ADAPTER arm_sensor (* Adapter Interface *)
  (* Standard: 61499-1 *)
  (* Version 0.0, 10/22/2026, lizar, Schneider Electric *)
  PACKAGE Main;
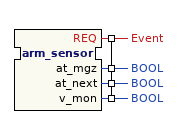
  EVENT_OUTPUT
    REQ WITH at_mgz, at_next, v_mon; (* Confirmation from Plug *)
  END_EVENT
  VAR_OUTPUT
    at_mgz : BOOL; (* Indication Data from Plug *)
    at_next : BOOL; (* Indication Data from Plug *)
    v_mon : BOOL; (* Indication Data from Plug *)
  END_VAR
  SERVICE SOCKET/PLUG
    SEQUENCE request_confirm
      SOCKET.REQ(REQD) -> PLUG.REQ(REQD);
      PLUG.REQ(CNFD) -> SOCKET.REQ(CNFD);
    END_SEQUENCE
    SEQUENCE indication_response
      PLUG.IND(at_mgz) -> SOCKET.IND(at_mgz);
      SOCKET.RSP(RSPD) -> PLUG.RSP(RSPD);
    END_SEQUENCE
  END_SERVICE
END_ADAPTER
